(* IEC 61131-3 sources: SRCI_CLIENT_PLC/RobotLibrary/Library/POUs/Additional/MC_WriteCallSubprogramCyclic/Structures, 2 files *)

(* ---- WriteCallSubprogramCyclicOutCmd.st ---- *)
{attribute 'pack_mode' := '1'}
// -------------------------------------------------------------------------
//  SRCI Robot Library
// -------------------------------------------------------------------------
//
//  Object:      UnitMeasurementOutCmd
//  Author:      Thorsten Brach
//  Date:        2024-08-11
//
//  Description:
//
//
//  Copyright:
//    (C) 2024 Thorsten Brach. All rights reserved
//             Licensed under the MIT License.
//
//  Disclaimer:
//    This project is provided without any guarantee and can be used for
//    private and commercial purposes. Any use is at the user’s
//    own risk and responsibility.
//
// -------------------------------------------------------------------------
TYPE WriteCallSubprogramCyclicOutCmd :
STRUCT

END_STRUCT
END_TYPE

(* ---- WriteCallSubprogramCyclicParCmd.st ---- *)
{attribute 'pack_mode' := '1'}
// -------------------------------------------------------------------------
//  SRCI Robot Library
// -------------------------------------------------------------------------
//
//  Object:      WriteCallSubprogramCyclicParCmd
//  Author:      Thorsten Brach
//  Date:        2024-08-11
//
//  Description:
//
//
//  Copyright:
//    (C) 2024 Thorsten Brach. All rights reserved
//             Licensed under the MIT License.
//
//  Disclaimer:
//    This project is provided without any guarantee and can be used for
//    private and commercial purposes. Any use is at the user’s
//    own risk and responsibility.
//
// -------------------------------------------------------------------------
TYPE WriteCallSubprogramCyclicParCmd :
STRUCT
  /// Cyclic input data of subprogram
  /// ST-FIX F179: size from RobotLibraryConstants.CYCLIC_SUB_PROGRAM_DATA_MAX
  Data : ARRAY[0..RobotLibraryConstants.CYCLIC_SUB_PROGRAM_DATA_MAX] OF BYTE;
END_STRUCT
END_TYPE
